Staubli VAL3: trajectory.pjx

--- trajectory.pjx ---
Parameters version=s8.15.3Cs9_BS3337 stackSize=5000 millimeterUnit=true
Program file=copy.pgx
Program file=copyPoint.pgx
Program file=copyPoint1.pgx
Program file=copyPoint3.pgx
Program file=deletePoint.pgx
Program file=deleteTraj.pgx
Program file=getFrameID.pgx
Program file=getIFvalue.pgx
Program file=getLibName.pgx
Program file=getMoveType.pgx
Program file=getPointIndex.pgx
Program file=getPointPara.pgx
Program file=getPointSize.pgx
Program file=getSize.pgx
Program file=getToolID.pgx
Program file=getTrajList.pgx
Program file=getTrajSize.pgx
Program file=insertAction.pgx
Program file=insertCirclePoint.pgx
Program file=insertDelay.pgx
Program file=insertENDIF.pgx
Program file=insertIF.pgx
Program file=insertJoint.pgx
Program file=insertPoint.pgx
Program file=insertSignal.pgx
Program file=isDefine.pgx
Program file=isPointOK.pgx
Program file=isReachable.pgx
Program file=loadTRAJ.pgx
Program file=logicIF.pgx
Program file=makeTraj.pgx
Program file=modifyAll.pgx
Program file=modifyPara.pgx
Program file=new.pgx
Program file=onSave.pgx
Program file=pointEdit.pgx
Program file=pointEditValue.pgx
Program file=pointMove.pgx
Program file=pointMove1.pgx
Program file=pointToString.pgx
Program file=resetMark.pgx
Program file=resizeMark.pgx
Program file=setMark.pgx
Program file=start.pgx
Program file=stop.pgx
Program file=teachPoint.pgx
Program file=teachPoint1.pgx
Data file=trajectory.dtx
Library alias=savedata path=Disk://source/saveData/saveData.pjx
Library alias=io path=Disk://source/projectSource/io/io.pjx
Library alias=rs path=Disk://source/projectSource/robotStatus/robotStatus.pjx
Library alias=actData path=Disk://data/actionData/actionData.pjx
Library alias=action path=Disk://source/projectSource/Action/Action.pjx
Library alias=trajTemp path=Disk://source/template/trajTemp/trajTemp.pjx
Library alias=ar path=Disk://autoReturn/autoReturn.pjx
Type name=pointItem path=Disk://source/template/pointItem/pointItem.pjx
Type name=trajItem path=Disk://source/template/trajItem/trajItem.pjx

--- trajectory.dtx ---
mdesc mNomSpeed
frame fFrame = {fatherId=world[0]}
tool tTool = {fatherId=flange[0]}
mdesc mSim = {blend=off}
frame _fFrame = {fatherId=world[0]}
pointRx pGOTO = {fatherId=world[0]}
num nIndex[100]

--- start.pgx ---
program start()
begin
end

--- copy.pgx ---
public program copy(string x_sSource, string& x_sTarget, bool& x_bToSave)
  local num l_j
  local num l_i
begin
  trajTemp:tTrajItem[x_sTarget].nFrameIndex=trajTemp:tTrajItem[x_sSource].nFrameIndex
  trajTemp:tTrajItem[x_sTarget].nToolIndex=trajTemp:tTrajItem[x_sSource].nToolIndex
  trajTemp:tTrajItem[x_sTarget].nMoveID=trajTemp:tTrajItem[x_sSource].nMoveID
  trajTemp:tTrajItem[x_sTarget].sID=trajTemp:tTrajItem[x_sTarget].sID
  resize(trajTemp:tTrajItem[x_sTarget].pPointItem,1,size(trajTemp:tTrajItem[x_sSource].pPointItem))
  for l_i = 0 to size(trajTemp:tTrajItem[x_sSource].pPointItem)-1
    trajTemp:tTrajItem[x_sTarget].pPointItem[l_i].pParaItem.mMdesc=trajTemp:tTrajItem[x_sSource].pPointItem[l_i].pParaItem.mMdesc
    trajTemp:tTrajItem[x_sTarget].pPointItem[l_i].pParaItem.nMoveType=trajTemp:tTrajItem[x_sSource].pPointItem[l_i].pParaItem.nMoveType
    trajTemp:tTrajItem[x_sTarget].pPointItem[l_i].pPointRx=trajTemp:tTrajItem[x_sSource].pPointItem[l_i].pPointRx
    //2025.03.18 add mlc  2025.10.16 modify by liu zhengang
    trajTemp:tTrajItem[x_sTarget].pPointItem[l_i].pInter=trajTemp:tTrajItem[x_sSource].pPointItem[l_i].pInter
    trajTemp:tTrajItem[x_sTarget].pPointItem[l_i].jJointRx=trajTemp:tTrajItem[x_sSource].pPointItem[l_i].jJointRx
    for l_j = 0 to 0
      trajTemp:tTrajItem[x_sTarget].pPointItem[l_i].pParaItem.nActionIndex[l_j]=trajTemp:tTrajItem[x_sSource].pPointItem[l_i].pParaItem.nActionIndex[l_j]
      trajTemp:tTrajItem[x_sTarget].pPointItem[l_i].pParaItem.nPercentage[l_j]=trajTemp:tTrajItem[x_sSource].pPointItem[l_i].pParaItem.nPercentage[l_j]
      trajTemp:tTrajItem[x_sTarget].pPointItem[l_i].pParaItem.iIfItem.bANDOR[l_j]=(trajTemp:tTrajItem[x_sSource].pPointItem[l_i].pParaItem.iIfItem.bANDOR[l_j]==true)
    endFor
    for l_j = 0 to 2
      trajTemp:tTrajItem[x_sTarget].pPointItem[l_i].pParaItem.iIfItem.nSigType[l_j]=trajTemp:tTrajItem[x_sSource].pPointItem[l_i].pParaItem.iIfItem.nSigType[l_j]
      trajTemp:tTrajItem[x_sTarget].pPointItem[l_i].pParaItem.iIfItem.nSigIndex[l_j]=trajTemp:tTrajItem[x_sSource].pPointItem[l_i].pParaItem.iIfItem.nSigIndex[l_j]
      trajTemp:tTrajItem[x_sTarget].pPointItem[l_i].pParaItem.iIfItem.nValue[l_j]=trajTemp:tTrajItem[x_sSource].pPointItem[l_i].pParaItem.iIfItem.nValue[l_j]
    endFor
    //
    trajTemp:tTrajItem[x_sTarget].pPointItem[l_i].pParaItem.nDelay=trajTemp:tTrajItem[x_sSource].pPointItem[l_i].pParaItem.nDelay
    trajTemp:tTrajItem[x_sTarget].pPointItem[l_i].pParaItem.nSigValue=trajTemp:tTrajItem[x_sSource].pPointItem[l_i].pParaItem.nSigValue
  endFor
  x_bToSave=true
end

--- copyPoint.pgx ---
public program copyPoint(string x_sKey, bool& x_bMark)
  local num l_nSize
  local num l_j
  local num l_i
begin
  resize(savedata:nMarkIndex,1,1)
  savedata:nMarkIndex=-1
  call getPointSize(x_sKey,l_nSize)
  l_j = 0
  for l_i = 0 to l_nSize-1
    if trajTemp:tTrajItem[x_sKey].pPointItem[l_i].bMarked
      l_j=l_j+1
      insert(savedata:nMarkIndex[l_j])
      savedata:nMarkIndex[l_j]=l_i


    endIf
  endFor
  x_bMark=false
end

--- copyPoint1.pgx ---
public program copyPoint1(string x_sKey, num x_nIndex)
  local num l_i
begin
  for l_i = 1 to size(savedata:nMarkIndex)-1
    insert(trajTemp:tTrajItem[x_sKey].pPointItem[x_nIndex+l_i])
    call copyPoint3(x_sKey,x_nIndex+l_i,savedata:nMarkIndex[l_i])
  endFor
  call resetMark(x_sKey)
end

--- copyPoint3.pgx ---
public program copyPoint3(string x_sKey, num x_nTarget, num x_nSource)
  local num l_i
begin
  trajTemp:tTrajItem[x_sKey].pPointItem[x_nTarget].pPointRx=trajTemp:tTrajItem[x_sKey].pPointItem[x_nSource].pPointRx
  //trajTemp:tTrajItem[x_sKey].pPointItem[x_nTarget].pPointRx[1]=trajTemp:tTrajItem[x_sKey].pPointItem[x_nSource].pPointRx[1]
  trajTemp:tTrajItem[x_sKey].pPointItem[x_nTarget].jJointRx=trajTemp:tTrajItem[x_sKey].pPointItem[x_nSource].jJointRx
  trajTemp:tTrajItem[x_sKey].pPointItem[x_nTarget].sID=trajTemp:tTrajItem[x_sKey].pPointItem[x_nSource].sID
  trajTemp:tTrajItem[x_sKey].pPointItem[x_nTarget].bMarked=trajTemp:tTrajItem[x_sKey].pPointItem[x_nSource].bMarked
  trajTemp:tTrajItem[x_sKey].pPointItem[x_nTarget].pInter=trajTemp:tTrajItem[x_sKey].pPointItem[x_nSource].pInter
  trajTemp:tTrajItem[x_sKey].pPointItem[x_nTarget].pParaItem.mMdesc=trajTemp:tTrajItem[x_sKey].pPointItem[x_nSource].pParaItem.mMdesc
  trajTemp:tTrajItem[x_sKey].pPointItem[x_nTarget].pParaItem.nMoveType=trajTemp:tTrajItem[x_sKey].pPointItem[x_nSource].pParaItem.nMoveType
  trajTemp:tTrajItem[x_sKey].pPointItem[x_nTarget].pParaItem.nActionIndex=trajTemp:tTrajItem[x_sKey].pPointItem[x_nSource].pParaItem.nActionIndex
  trajTemp:tTrajItem[x_sKey].pPointItem[x_nTarget].pParaItem.nPercentage=trajTemp:tTrajItem[x_sKey].pPointItem[x_nSource].pParaItem.nPercentage
  trajTemp:tTrajItem[x_sKey].pPointItem[x_nTarget].pParaItem.nDelay=trajTemp:tTrajItem[x_sKey].pPointItem[x_nSource].pParaItem.nDelay
  trajTemp:tTrajItem[x_sKey].pPointItem[x_nTarget].pParaItem.nSigValue=trajTemp:tTrajItem[x_sKey].pPointItem[x_nSource].pParaItem.nSigValue
  trajTemp:tTrajItem[x_sKey].pPointItem[x_nTarget].pParaItem.bSafePoint=trajTemp:tTrajItem[x_sKey].pPointItem[x_nSource].pParaItem.bSafePoint
  for l_i = 0 to 2
    trajTemp:tTrajItem[x_sKey].pPointItem[x_nTarget].pParaItem.iIfItem.nSigType[l_i]=trajTemp:tTrajItem[x_sKey].pPointItem[x_nSource].pParaItem.iIfItem.nSigType[l_i]
    trajTemp:tTrajItem[x_sKey].pPointItem[x_nTarget].pParaItem.iIfItem.nSigIndex[l_i]=trajTemp:tTrajItem[x_sKey].pPointItem[x_nSource].pParaItem.iIfItem.nSigIndex[l_i]
    trajTemp:tTrajItem[x_sKey].pPointItem[x_nTarget].pParaItem.iIfItem.nValue[l_i]=trajTemp:tTrajItem[x_sKey].pPointItem[x_nSource].pParaItem.iIfItem.nValue[l_i]
  endFor
  trajTemp:tTrajItem[x_sKey].pPointItem[x_nTarget].pParaItem.iIfItem.bANDOR[0]=trajTemp:tTrajItem[x_sKey].pPointItem[x_nSource].pParaItem.iIfItem.bANDOR[0]
  trajTemp:tTrajItem[x_sKey].pPointItem[x_nTarget].pParaItem.iIfItem.bANDOR[1]=trajTemp:tTrajItem[x_sKey].pPointItem[x_nSource].pParaItem.iIfItem.bANDOR[1]

end

--- deletePoint.pgx ---
public program deletePoint(string x_sKey, num x_nIndex, bool& x_bToSave)
  local bool l_bResult
begin
  l_bResult=userPageConfirm("是否删除点位："+toString("",x_nIndex))
  if l_bResult
    if x_nIndex==0 and size(trajTemp:tTrajItem[x_sKey].pPointItem)==1
      userPageAlert("数组元素不得为0")
    else
      delete(trajTemp:tTrajItem[x_sKey].pPointItem[x_nIndex])
      //trajTemp:libSave()
      x_bToSave=true
    endIf
  endIf

end

--- deleteTraj.pgx ---
public program deleteTraj(string x_sKey, bool& x_bToSave)
begin
  if isDefined(trajTemp:tTrajItem[x_sKey])
    delete(trajTemp:tTrajItem[x_sKey])
    //trajTemp:libSave()
  endIf
  x_bToSave=true
end

--- getFrameID.pgx ---
public program getFrameID(string x_sKey, num& x_nFrameID)
begin
  x_nFrameID=trajTemp:tTrajItem[x_sKey].nFrameIndex
end

--- getIFvalue.pgx ---
public program getIFvalue(string x_sKey, num x_nIndex, bool& x_bFinalResult)
  local num l_nSigType[3]
  local num l_i
  local num l_nSigValue[3]
  local bool l_bANDOR[2]
  local num l_nSigIndex[3]
  local bool l_bValue
  local bool l_bErr
  local bool l_bSetValue
  local num l_nResult[3]
  local bool l_bResult0[2]
  local num l_nValue
begin
  //l_nResult=0,null
  //         =1,true
  //         =2,false

  for l_i = 0 to 2
    l_nSigType[l_i]= trajTemp:tTrajItem[x_sKey].pPointItem[x_nIndex].pParaItem.iIfItem.nSigType[l_i]
    l_nSigValue[l_i]=trajTemp:tTrajItem[x_sKey].pPointItem[x_nIndex].pParaItem.iIfItem.nValue[l_i]
    l_nSigIndex[l_i]=trajTemp:tTrajItem[x_sKey].pPointItem[x_nIndex].pParaItem.iIfItem.nSigIndex[l_i]
  endFor
  l_bANDOR[0]=trajTemp:tTrajItem[x_sKey].pPointItem[x_nIndex].pParaItem.iIfItem.bANDOR[0]
  l_bANDOR[1]=trajTemp:tTrajItem[x_sKey].pPointItem[x_nIndex].pParaItem.iIfItem.bANDOR[1]

  for l_i = 0 to 2
    if l_nSigType[l_i]!=0 and l_nSigIndex[l_i]!=0
      switch l_nSigType[l_i]
        case 1
          //din
          call io:getDigIO(io:dInput[l_nSigIndex[l_i]],l_bValue,l_bErr)
          l_bSetValue=(l_nSigValue[l_i]!=0)
          if l_bSetValue==l_bValue
            l_nResult[l_i]=1
          else
            l_nResult[l_i]=2
          endIf
        break
        case 2
          //dout
          call io:getDigIO(io:dOutput[l_nSigIndex[l_i]],l_bValue,l_bErr)
          l_bSetValue=(l_nSigValue[l_i]!=0)
          if l_bSetValue==l_bValue
            l_nResult[l_i]=1
          else
            l_nResult[l_i]=2
          endIf
        break
        case 3
          //ain
          call io:getAnaIO(io:aInput[l_nSigIndex[l_i]],l_nValue,l_bErr)
          if l_nSigValue[l_i]==l_nValue
            l_nResult[l_i]=1
          else
            l_nResult[l_i]=2
          endIf
        break
        case 4
          //aout
          call io:getAnaIO(io:aOutput[l_nSigIndex[l_i]],l_nValue,l_bErr)
          if l_nSigValue[l_i]==l_nValue
            l_nResult[l_i]=1
          else
            l_nResult[l_i]=2
          endIf
        break
      endSwitch
    else
      l_nResult[l_i]=0
    endIf
  endFor

  //logic
 call logicIF(l_nResult[0],l_nResult[1],l_nResult[2],l_bANDOR[0],l_bANDOR[1],x_bFinalResult)

end

--- getLibName.pgx ---
public program getLibName(num& x_nLibNum, bool& x_bResult)
  local string l_sString
  local string l_sString1
  local num l_nPos
  local string l_sPath
  local num l_nlength
  local num l_nlength1
  local num l_nLength2
  local num l_nSize
  local string l_sTarget
  local num l_nLength
begin
  l_sPath=trajTemp:libPath()
  l_nlength=len("Disk://data/CustomerLib/lib")
  l_nlength1=len("/saveTRAJ/saveTRAJ.pjx")
  l_nLength2=len(l_sPath)
  l_nSize=l_nLength2-l_nlength1-l_nLength
  l_sTarget=mid(l_sPath,l_nSize,l_nlength)
  toNum(l_sTarget,x_nLibNum,x_bResult)
end

--- getMoveType.pgx ---
public program getMoveType(string x_sKey, num x_nIndex, num& x_nMoveType)
begin
  x_nMoveType=trajTemp:tTrajItem[x_sKey].pPointItem[x_nIndex].pParaItem.nMoveType
end

--- getPointIndex.pgx ---
public program getPointIndex(string x_sTrajItem, string x_sPoint, num& x_nPointIndex, bool& x_bResult)
  local bool l_bResult
  local num l_nSize
begin
  toNum(x_sPoint,x_nPointIndex,x_bResult)
  if !x_bResult
    call getPointSize(x_sTrajItem,l_nSize)
    x_nPointIndex=l_nSize-1
  endIf
end

--- getPointPara.pgx ---
public program getPointPara(string x_sKey, num x_nIndex, num& x_nMoveType, num& x_nParaSpeed, num& x_nParaAccel, num& x_nParaBlend, num x_nParaPercent, string& x_sComment, bool& x_bSafePoint, string& x_sBlend, num& x_nValue[], string& x_sTRSF[])
  local num l_nMoveType
begin
  x_nMoveType=trajTemp:tTrajItem[x_sKey].pPointItem[x_nIndex].pParaItem.nMoveType
  x_nParaSpeed=trajTemp:tTrajItem[x_sKey].pPointItem[x_nIndex].pParaItem.mMdesc.vel
  x_nParaAccel=trajTemp:tTrajItem[x_sKey].pPointItem[x_nIndex].pParaItem.mMdesc.accel
  x_nParaBlend=trajTemp:tTrajItem[x_sKey].pPointItem[x_nIndex].pParaItem.mMdesc.leave
  x_nParaPercent=trajTemp:tTrajItem[x_sKey].pPointItem[x_nIndex].pParaItem.nPercentage
  x_sComment=trajTemp:tTrajItem[x_sKey].pPointItem[x_nIndex].sID
  //  x_bBlendJoint=(trajTemp:tTrajItem[x_sKey].pPointItem[x_nIndex].pParaItem.mMdesc.blend==joint)
  //  x_bBlendOFF=(trajTemp:tTrajItem[x_sKey].pPointItem[x_nIndex].pParaItem.mMdesc.blend==off)
  switch x_nMoveType
    case 1

      x_nValue[0]=trajTemp:tTrajItem[x_sKey].pPointItem[x_nIndex].jJointRx.j1
      x_nValue[1]=trajTemp:tTrajItem[x_sKey].pPointItem[x_nIndex].jJointRx.j2
      x_nValue[2]=trajTemp:tTrajItem[x_sKey].pPointItem[x_nIndex].jJointRx.j3
      x_nValue[3]=trajTemp:tTrajItem[x_sKey].pPointItem[x_nIndex].jJointRx.j4
      x_nValue[4]=trajTemp:tTrajItem[x_sKey].pPointItem[x_nIndex].jJointRx.j5
      x_nValue[5]=trajTemp:tTrajItem[x_sKey].pPointItem[x_nIndex].jJointRx.j6

      x_sTRSF[0]="J1:"
      x_sTRSF[1]="J2:"
      x_sTRSF[2]="J3:"
      x_sTRSF[3]="J4:"
      x_sTRSF[4]="J5:"
      x_sTRSF[5]="J6:"

    break
    case 0
      x_nValue[0]=trajTemp:tTrajItem[x_sKey].pPointItem[x_nIndex].pPointRx.trsf.x
      x_nValue[1]=trajTemp:tTrajItem[x_sKey].pPointItem[x_nIndex].pPointRx.trsf.y
      x_nValue[2]=trajTemp:tTrajItem[x_sKey].pPointItem[x_nIndex].pPointRx.trsf.z
      x_nValue[3]=trajTemp:tTrajItem[x_sKey].pPointItem[x_nIndex].pPointRx.trsf.rx
      x_nValue[4]=trajTemp:tTrajItem[x_sKey].pPointItem[x_nIndex].pPointRx.trsf.ry
      x_nValue[5]=trajTemp:tTrajItem[x_sKey].pPointItem[x_nIndex].pPointRx.trsf.rz

      x_sTRSF[0]="X:"
      x_sTRSF[1]="Y:"
      x_sTRSF[2]="Z:"
      x_sTRSF[3]="RX:"
      x_sTRSF[4]="RY:"
      x_sTRSF[5]="RZ:"
    break
    case 2
      x_nValue[0]=trajTemp:tTrajItem[x_sKey].pPointItem[x_nIndex].pPointRx.trsf.x
      x_nValue[1]=trajTemp:tTrajItem[x_sKey].pPointItem[x_nIndex].pPointRx.trsf.y
      x_nValue[2]=trajTemp:tTrajItem[x_sKey].pPointItem[x_nIndex].pPointRx.trsf.z
      x_nValue[3]=trajTemp:tTrajItem[x_sKey].pPointItem[x_nIndex].pPointRx.trsf.rx
      x_nValue[4]=trajTemp:tTrajItem[x_sKey].pPointItem[x_nIndex].pPointRx.trsf.ry
      x_nValue[5]=trajTemp:tTrajItem[x_sKey].pPointItem[x_nIndex].pPointRx.trsf.rz
      x_nValue[6]= trajTemp:tTrajItem[x_sKey].pPointItem[x_nIndex].pInter.trsf.x
      x_nValue[7]=trajTemp:tTrajItem[x_sKey].pPointItem[x_nIndex].pInter.trsf.y
      x_nValue[8]=trajTemp:tTrajItem[x_sKey].pPointItem[x_nIndex].pInter.trsf.z
      x_nValue[9]=trajTemp:tTrajItem[x_sKey].pPointItem[x_nIndex].pInter.trsf.rx
      x_nValue[10]=trajTemp:tTrajItem[x_sKey].pPointItem[x_nIndex].pInter.trsf.ry
      x_nValue[11]= trajTemp:tTrajItem[x_sKey].pPointItem[x_nIndex].pInter.trsf.rz
      x_sTRSF[0]="X:"
      x_sTRSF[1]="Y:"
      x_sTRSF[2]="Z:"
      x_sTRSF[3]="RX:"
      x_sTRSF[4]="RY:"
      x_sTRSF[5]="RZ:"
      x_sTRSF[6]="2X:"
      x_sTRSF[7]="2Y:"
      x_sTRSF[8]="2Z:"
      x_sTRSF[9]="2RX:"
      x_sTRSF[10]="2RY:"
      x_sTRSF[11]="2RZ:"

    break
  endSwitch
  //blend
  if trajTemp:tTrajItem[x_sKey].pPointItem[x_nIndex].pParaItem.mMdesc.blend==off
    x_sBlend="OFF"
  elseIf trajTemp:tTrajItem[x_sKey].pPointItem[x_nIndex].pParaItem.mMdesc.blend==joint
    x_sBlend="关节"
  elseIf trajTemp:tTrajItem[x_sKey].pPointItem[x_nIndex].pParaItem.mMdesc.blend==Cartesian
    x_sBlend="笛卡尔"
  endIf
  x_bSafePoint = (trajTemp:tTrajItem[x_sKey].pPointItem.pParaItem.bSafePoint==true)
end

--- getPointSize.pgx ---
public program getPointSize(string x_sKey, num& x_nSize)
begin
  x_nSize=size(trajTemp:tTrajItem[x_sKey].pPointItem)
end

--- getSize.pgx ---
public program getSize(num& x_nSize)
begin
  if size(trajTemp:tTrajItem)>0
    x_nSize=size(trajTemp:tTrajItem)
  else
    x_nSize=0
  endIf
end

--- getToolID.pgx ---
public program getToolID(string x_sKey, num& x_nToolID)
begin
   x_nToolID=trajTemp:tTrajItem[x_sKey].nToolIndex
end

--- getTrajList.pgx ---
public program getTrajList(string& x_sList[])
  local string l_sKey
begin
  resize(x_sList,1,1)
  l_sKey=first(trajTemp:tTrajItem)

  while l_sKey!=""
    x_sList[size(x_sList)-1]=l_sKey

    l_sKey=next(trajTemp:tTrajItem[l_sKey])

    if l_sKey!=""
      insert(x_sList[size(x_sList)])
    endIf
  endWhile
  if size(trajTemp:tTrajItem)<1
    x_sList=""
  endIf
end

--- getTrajSize.pgx ---
public program getTrajSize(num& x_nSize)
begin
  x_nSize=size(trajTemp:tTrajItem)
end

--- insertAction.pgx ---
public program insertAction(string x_sKey, num x_nIndex, num x_nValue, bool& x_bToSave)
  local num l_i
begin
  // insert(trajTemp:tTrajItem[x_sKey].pPointItem[x_nIndex+1])
  append(trajTemp:tTrajItem[x_sKey].pPointItem)

  for l_i = (size(trajTemp:tTrajItem[x_sKey].pPointItem)-1) to(x_nIndex+1) step -1
    //logMsg(toString("",l_i))
    call copyPoint3(x_sKey,l_i,l_i-1)
  endFor
  trajTemp:tTrajItem[x_sKey].pPointItem[x_nIndex+1].pParaItem.nMoveType=10
  trajTemp:tTrajItem[x_sKey].pPointItem[x_nIndex+1].pParaItem.nSigValue=x_nValue
  //trajTemp:libSave()
  x_bToSave=true
end

--- insertCirclePoint.pgx ---
public program insertCirclePoint(string x_sKey, num x_nIndex, bool& x_bToSave)
  local num l_j
  local frame l_fFrame
  local tool l_tTool
  local num l_i
  local num l_nFrameIndex
  local num l_nToolIndex
  local pointRx l_pPoint
begin
  //  link(l_fFrame,world)
  //  link(l_tTool,flange)
  //  call savedata:getFrame(trajTemp:tTrajItem[x_sKey].nFrameIndex,l_fFrame)
  //  call savedata:getTool(trajTemp:tTrajItem[x_sKey].nToolIndex,l_tTool)
  //insert(trajTemp:tTrajItem[x_sKey].pPointItem[x_nIndex+1])
  append(trajTemp:tTrajItem[x_sKey].pPointItem)

  for l_i = (size(trajTemp:tTrajItem[x_sKey].pPointItem)-1) to(x_nIndex+1) step -1
    //logMsg(toString("",l_i))
    call copyPoint3(x_sKey,l_i,l_i-1)
  endFor
  //2024.12.06 当前位置作为插入点坐标
  l_nFrameIndex=trajTemp:tTrajItem[x_sKey].nFrameIndex
  l_nToolIndex=trajTemp:tTrajItem[x_sKey].nToolIndex
  call savedata:getFrame(l_nFrameIndex,l_fFrame)
  call savedata:getTool(l_nToolIndex,l_tTool)
  trajTemp:tTrajItem[x_sKey].pPointItem[x_nIndex+1].jJointRx=herej()
  l_pPoint=jointToPoint(l_tTool,l_fFrame,herej())
  trajTemp:tTrajItem[x_sKey].pPointItem[x_nIndex+1].pPointRx.trsf=l_pPoint.trsf
  trajTemp:tTrajItem[x_sKey].pPointItem[x_nIndex+1].pPointRx.config=l_pPoint.config
  trajTemp:tTrajItem[x_sKey].pPointItem[x_nIndex+1].pInter.trsf=l_pPoint.trsf
  trajTemp:tTrajItem[x_sKey].pPointItem[x_nIndex+1].pInter.config=l_pPoint.config
  //

  //trajTemp:tTrajItem[x_sKey].pPointItem[x_nIndex+1].pPointRx=trajTemp:tTrajItem[x_sKey].pPointItem[x_nIndex].pPointRx
  //trajTemp:tTrajItem[x_sKey].pPointItem[x_nIndex+1].jJointRx=trajTemp:tTrajItem[x_sKey].pPointItem[x_nIndex].jJointRx
  trajTemp:tTrajItem[x_sKey].pPointItem[x_nIndex+1].pParaItem.mMdesc=trajTemp:tTrajItem[x_sKey].pPointItem[x_nIndex].pParaItem.mMdesc
  trajTemp:tTrajItem[x_sKey].pPointItem[x_nIndex+1].pParaItem.nMoveType=2
  trajTemp:tTrajItem[x_sKey].pPointItem[x_nIndex+1].pParaItem.nDelay=trajTemp:tTrajItem[x_sKey].pPointItem[x_nIndex].pParaItem.nDelay
  trajTemp:tTrajItem[x_sKey].pPointItem[x_nIndex+1].pParaItem.nSigValue=trajTemp:tTrajItem[x_sKey].pPointItem[x_nIndex].pParaItem.nSigValue
  trajTemp:tTrajItem[x_sKey].pPointItem[x_nIndex+1].pParaItem.nActionIndex=trajTemp:tTrajItem[x_sKey].pPointItem[x_nIndex].pParaItem.nActionIndex
  trajTemp:tTrajItem[x_sKey].pPointItem[x_nIndex+1].pParaItem.nPercentage=trajTemp:tTrajItem[x_sKey].pPointItem[x_nIndex].pParaItem.nPercentage
  for l_j = 0 to 2
    trajTemp:tTrajItem[x_sKey].pPointItem[x_nIndex+1].pParaItem.iIfItem.nSigType[l_j]=trajTemp:tTrajItem[x_sKey].pPointItem[x_nIndex].pParaItem.iIfItem.nSigType[l_j]
    trajTemp:tTrajItem[x_sKey].pPointItem[x_nIndex+1].pParaItem.iIfItem.nSigIndex[l_j]=trajTemp:tTrajItem[x_sKey].pPointItem[x_nIndex].pParaItem.iIfItem.nSigIndex[l_j]
    trajTemp:tTrajItem[x_sKey].pPointItem[x_nIndex+1].pParaItem.iIfItem.nValue[l_j]=trajTemp:tTrajItem[x_sKey].pPointItem[x_nIndex].pParaItem.iIfItem.nValue[l_j]
  endFor
  //trajTemp:libSave()
  x_bToSave=true
end

--- insertDelay.pgx ---
public program insertDelay(string x_sKey, num x_nIndex, bool& x_bToSave, num x_nMoveType, num x_nDelay)
  local num l_j
  local num l_i
begin
  //insert(trajTemp:tTrajItem[x_sKey].pPointItem[x_nIndex+1])
  append(trajTemp:tTrajItem[x_sKey].pPointItem)

  for l_i = (size(trajTemp:tTrajItem[x_sKey].pPointItem)-1) to(x_nIndex+1) step -1
   // logMsg(toString("",l_i))
    call copyPoint3(x_sKey,l_i,l_i-1)
  endFor
  trajTemp:tTrajItem[x_sKey].pPointItem[x_nIndex+1].pParaItem.nMoveType=x_nMoveType

  trajTemp:tTrajItem[x_sKey].pPointItem[x_nIndex+1].pParaItem.nDelay=x_nDelay

 //trajTemp:libSave()

  x_bToSave=true
end

--- insertENDIF.pgx ---
public program insertENDIF(string x_sKey, num x_nIndex, bool& x_bToSave)
  local num l_j
  local num l_i
begin

  //insert(trajTemp:tTrajItem[x_sKey].pPointItem[x_nIndex+1])
  append(trajTemp:tTrajItem[x_sKey].pPointItem)

  for l_i = (size(trajTemp:tTrajItem[x_sKey].pPointItem)-1) to(x_nIndex+1) step -1
    //logMsg(toString("",l_i))
    call copyPoint3(x_sKey,l_i,l_i-1)
  endFor
  trajTemp:tTrajItem[x_sKey].pPointItem[x_nIndex+1].pParaItem.nMoveType=9

  //trajTemp:libSave()
  x_bToSave=true
end

--- insertIF.pgx ---
public program insertIF(string x_sKey, num x_nIndex, num& x_nMoveType[], num& x_nIOIndex[], num& x_nValue[], num& x_nANDOR[], bool& x_bToSave)
  local num l_j
  local num l_i
begin
  // insert(trajTemp:tTrajItem[x_sKey].pPointItem[x_nIndex+1])
  append(trajTemp:tTrajItem[x_sKey].pPointItem)

  for l_i = (size(trajTemp:tTrajItem[x_sKey].pPointItem)-1) to(x_nIndex+1) step -1
    // logMsg(toString("",l_i))
    call copyPoint3(x_sKey,l_i,l_i-1)
  endFor
  trajTemp:tTrajItem[x_sKey].pPointItem[x_nIndex+1].pParaItem.nMoveType=8
  for l_i =0 to 2
    trajTemp:tTrajItem[x_sKey].pPointItem[x_nIndex+1].pParaItem.iIfItem.nSigType[l_i]=x_nMoveType[l_i]
    trajTemp:tTrajItem[x_sKey].pPointItem[x_nIndex+1].pParaItem.iIfItem.nSigIndex[l_i]=x_nIOIndex[l_i]
    trajTemp:tTrajItem[x_sKey].pPointItem[x_nIndex+1].pParaItem.iIfItem.nValue[l_i]=x_nValue[l_i]
  endFor
  for l_i = 0 to 1
    trajTemp:tTrajItem[x_sKey].pPointItem[x_nIndex+1].pParaItem.iIfItem.bANDOR[l_i]=(x_nANDOR[l_i]==2)
  endFor

  //trajTemp:libSave()
  x_bToSave=true
end

--- insertJoint.pgx ---
public program insertJoint(string x_sKey, num x_nIndex, bool& x_bToSave)
  local num l_j
  local num l_i
begin
  // insert(trajTemp:tTrajItem[x_sKey].pPointItem[x_nIndex+1])
  append(trajTemp:tTrajItem[x_sKey].pPointItem)

  for l_i = (size(trajTemp:tTrajItem[x_sKey].pPointItem)-1) to(x_nIndex+1) step -1
    //logMsg(toString("",l_i))
    call copyPoint3(x_sKey,l_i,l_i-1)
  endFor
  trajTemp:tTrajItem[x_sKey].pPointItem[x_nIndex+1].pPointRx=trajTemp:tTrajItem[x_sKey].pPointItem[x_nIndex].pPointRx
  trajTemp:tTrajItem[x_sKey].pPointItem[x_nIndex+1].jJointRx=trajTemp:tTrajItem[x_sKey].pPointItem[x_nIndex].jJointRx
  trajTemp:tTrajItem[x_sKey].pPointItem[x_nIndex+1].pParaItem.mMdesc=trajTemp:tTrajItem[x_sKey].pPointItem[x_nIndex].pParaItem.mMdesc
  trajTemp:tTrajItem[x_sKey].pPointItem[x_nIndex+1].pParaItem.nMoveType=0
  trajTemp:tTrajItem[x_sKey].pPointItem[x_nIndex+1].pParaItem.nDelay=trajTemp:tTrajItem[x_sKey].pPointItem[x_nIndex].pParaItem.nDelay
  trajTemp:tTrajItem[x_sKey].pPointItem[x_nIndex+1].pParaItem.nSigValue=trajTemp:tTrajItem[x_sKey].pPointItem[x_nIndex].pParaItem.nSigValue
  trajTemp:tTrajItem[x_sKey].pPointItem[x_nIndex+1].pParaItem.nActionIndex=trajTemp:tTrajItem[x_sKey].pPointItem[x_nIndex].pParaItem.nActionIndex
  trajTemp:tTrajItem[x_sKey].pPointItem[x_nIndex+1].pParaItem.nPercentage=trajTemp:tTrajItem[x_sKey].pPointItem[x_nIndex].pParaItem.nPercentage
  for l_j = 0 to 2
    trajTemp:tTrajItem[x_sKey].pPointItem[x_nIndex+1].pParaItem.iIfItem.nSigType[l_j]=trajTemp:tTrajItem[x_sKey].pPointItem[x_nIndex].pParaItem.iIfItem.nSigType[l_j]
    trajTemp:tTrajItem[x_sKey].pPointItem[x_nIndex+1].pParaItem.iIfItem.nSigIndex[l_j]=trajTemp:tTrajItem[x_sKey].pPointItem[x_nIndex].pParaItem.iIfItem.nSigIndex[l_j]
    trajTemp:tTrajItem[x_sKey].pPointItem[x_nIndex+1].pParaItem.iIfItem.nValue[l_j]=trajTemp:tTrajItem[x_sKey].pPointItem[x_nIndex].pParaItem.iIfItem.nValue[l_j]
  endFor
  //trajTemp:libSave()
  x_bToSave=true
end

--- insertPoint.pgx ---
public program insertPoint(string x_sKey, num x_nIndex, bool& x_bToSave)
  local num l_j
  local frame l_fFrame
  local tool l_tTool
  local num l_i
begin
  //  link(l_fFrame,world)
  //  link(l_tTool,flange)
  //  call savedata:getFrame(trajTemp:tTrajItem[x_sKey].nFrameIndex,l_fFrame)
  //  call savedata:getTool(trajTemp:tTrajItem[x_sKey].nToolIndex,l_tTool)
  //insert(trajTemp:tTrajItem[x_sKey].pPointItem[x_nIndex+1])
   append(trajTemp:tTrajItem[x_sKey].pPointItem)

  for l_i = (size(trajTemp:tTrajItem[x_sKey].pPointItem)-1) to(x_nIndex+1) step -1
    //logMsg(toString("",l_i))
    call copyPoint3(x_sKey,l_i,l_i-1)
  endFor
  trajTemp:tTrajItem[x_sKey].pPointItem[x_nIndex+1].pPointRx=trajTemp:tTrajItem[x_sKey].pPointItem[x_nIndex].pPointRx
  trajTemp:tTrajItem[x_sKey].pPointItem[x_nIndex+1].jJointRx=trajTemp:tTrajItem[x_sKey].pPointItem[x_nIndex].jJointRx
  trajTemp:tTrajItem[x_sKey].pPointItem[x_nIndex+1].pParaItem.mMdesc=trajTemp:tTrajItem[x_sKey].pPointItem[x_nIndex].pParaItem.mMdesc
  trajTemp:tTrajItem[x_sKey].pPointItem[x_nIndex+1].pParaItem.nMoveType=1
  trajTemp:tTrajItem[x_sKey].pPointItem[x_nIndex+1].pParaItem.nDelay=trajTemp:tTrajItem[x_sKey].pPointItem[x_nIndex].pParaItem.nDelay
  trajTemp:tTrajItem[x_sKey].pPointItem[x_nIndex+1].pParaItem.nSigValue=trajTemp:tTrajItem[x_sKey].pPointItem[x_nIndex].pParaItem.nSigValue
  trajTemp:tTrajItem[x_sKey].pPointItem[x_nIndex+1].pParaItem.nActionIndex=trajTemp:tTrajItem[x_sKey].pPointItem[x_nIndex].pParaItem.nActionIndex
  trajTemp:tTrajItem[x_sKey].pPointItem[x_nIndex+1].pParaItem.nPercentage=trajTemp:tTrajItem[x_sKey].pPointItem[x_nIndex].pParaItem.nPercentage
  for l_j = 0 to 2
    trajTemp:tTrajItem[x_sKey].pPointItem[x_nIndex+1].pParaItem.iIfItem.nSigType[l_j]=trajTemp:tTrajItem[x_sKey].pPointItem[x_nIndex].pParaItem.iIfItem.nSigType[l_j]
    trajTemp:tTrajItem[x_sKey].pPointItem[x_nIndex+1].pParaItem.iIfItem.nSigIndex[l_j]=trajTemp:tTrajItem[x_sKey].pPointItem[x_nIndex].pParaItem.iIfItem.nSigIndex[l_j]
    trajTemp:tTrajItem[x_sKey].pPointItem[x_nIndex+1].pParaItem.iIfItem.nValue[l_j]=trajTemp:tTrajItem[x_sKey].pPointItem[x_nIndex].pParaItem.iIfItem.nValue[l_j]
  endFor
  //trajTemp:libSave()
  x_bToSave=true
end

--- insertSignal.pgx ---
public program insertSignal(string x_sKey, num x_nIndex, bool& x_bToSave, num x_nMoveType, num x_nActionIndex, num x_nSigValue)
  local num l_j
  local bool l_bResult
  local num l_nIndex
  local num l_i
begin
  l_nIndex=x_nIndex+1

  //insert(trajTemp:tTrajItem[x_sKey].pPointItem[l_nIndex])
  append(trajTemp:tTrajItem[x_sKey].pPointItem)

  for l_i = (size(trajTemp:tTrajItem[x_sKey].pPointItem)-1) to l_nIndex step -1
    // logMsg(toString("",l_i))
    call copyPoint3(x_sKey,l_i,l_i-1)
  endFor
  trajTemp:tTrajItem[x_sKey].pPointItem[l_nIndex].pParaItem.nMoveType=x_nMoveType

  trajTemp:tTrajItem[x_sKey].pPointItem[l_nIndex].pParaItem.nSigValue=x_nSigValue

  trajTemp:tTrajItem[x_sKey].pPointItem[l_nIndex].pParaItem.nActionIndex=x_nActionIndex



  x_bToSave=true
  //trajTemp:libSave()
end

--- isDefine.pgx ---
public program isDefine(string x_sKey, bool& x_bResult)
begin
  x_bResult=isDefined(trajTemp:tTrajItem[x_sKey])
end

--- isPointOK.pgx ---
public program isPointOK(string x_sKey, num x_nIndex, bool& x_bResult)
  local pointRx l_pPoint
  local num l_nToolID
  local tool l_tTool
  local frame l_fFrame
  local num l_nFrameID
  local bool l_bResult
  local jointRx l_jResult
begin
  link(l_tTool,flange)
  link(l_fFrame,world)
  call getFrameID(x_sKey,l_nFrameID)
  call getToolID(x_sKey,l_nToolID)
  call savedata:getTool(l_nToolID,l_tTool)
  call savedata:getFrame(l_nFrameID,l_fFrame)
  link(l_pPoint,l_fFrame)
  l_pPoint.trsf=trajTemp:tTrajItem[x_sKey].pPointItem[x_nIndex].pPointRx.trsf
  l_pPoint.config=trajTemp:tTrajItem[x_sKey].pPointItem[x_nIndex].pPointRx.config

  l_bResult=pointToJoint(l_tTool,herej(),l_pPoint,l_jResult)
  if l_pPoint.trsf!={0,0,0,0,0,0} and l_bResult and isInRange(l_jResult)
    x_bResult=true
  else
    x_bResult=false
  endIf
end

--- isReachable.pgx ---
public program isReachable(string x_sKey, num x_nIndex, tool x_tTool)
  local pointRx l_pPoint
  local bool l_bResult
  local mdesc l_mDesc
  local jointRx l_jJoint
begin
  if trajTemp:tTrajItem[x_sKey].pPointItem[x_nIndex].pParaItem.nMoveType==0
    l_mDesc=trajTemp:tTrajItem[x_sKey].pPointItem[x_nIndex].pParaItem.mMdesc
    l_pPoint.trsf=trajTemp:tTrajItem[x_sKey].pPointItem.pPointRx.trsf
    l_pPoint.config=trajTemp:tTrajItem[x_sKey].pPointItem.pPointRx.config
    l_bResult= pointToJoint(x_tTool,herej(),l_pPoint,l_jJoint)
    if l_bResult
      movel(l_pPoint,x_tTool,l_mDesc)
    endIf
  endIf
end

--- loadTRAJ.pgx ---
public program loadTRAJ(num x_nLib, num& x_nResult)
  local string l_sPath
  local num l_nResult
begin
  if x_nLib>=0
    l_sPath="Disk://data/CustomerLib/lib"+toString("",x_nLib)+"/saveTRAJ"
    //  if libList()
    //    endIf
    x_nResult=trajTemp:libLoad(l_sPath)
    if x_nResult!=0
      popUpMsg("2")
      call rs:setAlarm(300,0)
    endIf
  else
    call rs:setAlarm(302,0)
  endIf
end

--- logicIF.pgx ---
public program logicIF(num x_nResult1, num x_nResult2, num x_nResult3, bool x_bANDOR1, bool x_bANDOR2, bool& x_bFinalResult)
  local bool l_bFinalResult1
  local bool l_bFinalResult2
begin
  if x_nResult1==0 and x_nResult2==0 and x_nResult3==0
    x_bFinalResult=false
  elseIf x_nResult1==0 and x_nResult2==0 and x_nResult3!=0
    x_bFinalResult=(x_nResult3==1)
  elseIf x_nResult1==0 and x_nResult2!=0 and x_nResult3==0
    x_bFinalResult=(x_nResult2==1)
  elseIf x_nResult1!=0 and x_nResult2==0 and x_nResult3==0
    x_bFinalResult=(x_nResult1==1)
  elseIf x_nResult1!=0 and x_nResult2!=0 and x_nResult3==0
    if x_bANDOR1
      x_bFinalResult=(x_nResult1==1 or x_nResult2==1)
    else
      x_bFinalResult=(x_nResult1==1 and x_nResult2==1)
    endIf
  elseIf x_nResult1==0 and x_nResult2!=0 and x_nResult3!=0
    if x_bANDOR2
      x_bFinalResult=(x_nResult1==1 or x_nResult2==1)
    else
      x_bFinalResult=(x_nResult1==1 and x_nResult2==1)
    endIf
  elseIf x_nResult1!=0 and x_nResult2!=0 and x_nResult3!=0
    if x_bANDOR1 and x_bANDOR2
      x_bFinalResult=(x_nResult1==1 or x_nResult2==1 or x_nResult3==1)
    elseIf !x_bANDOR1 and !x_bANDOR2
      x_bFinalResult=(x_nResult1==1 and x_nResult2==1 and x_nResult3==1)
    elseIf !x_bANDOR1 and x_bANDOR2
      x_bFinalResult=(x_nResult1==1 and x_nResult2==1 or x_nResult3==1)
    elseIf x_bANDOR1 and !x_bANDOR2
      x_bFinalResult=((x_nResult1==1 or x_nResult2==1) and x_nResult3==1)
    endIf

  endIf
end

--- makeTraj.pgx ---
public program makeTraj(string x_sKey)
  local num l_nMoveType
  local num l_nMoveID
  local frame l_fFrame
  local tool l_tTool
  local pointRx l_pPoint[2]
  local jointRx l_jJoint
  local mdesc l_mDesc
  local num l_nSigIndex
  local num l_nValue
  local bool l_bErr
  local num l_nSigValue
  local bool l_bValue
  local bool l_bSigValue
  local num l_i
  local num l_nDelay
  local bool l_bResult
  local num l_nActIndex
  local num l_nGetID
  local string l_sMsg
begin
  rs:sTrajStatus="执行轨迹："+x_sKey
  rs:sCycleItem=x_sKey
  l_nMoveID=trajTemp:tTrajItem[x_sKey].nMoveID
  rs:nFrameIndex=trajTemp:tTrajItem[x_sKey].nFrameIndex
  rs:nToolIndex=trajTemp:tTrajItem[x_sKey].nToolIndex
  call savedata:getFrame(rs:nFrameIndex,l_fFrame)
  call savedata:getTool(rs:nToolIndex,l_tTool)
  waitEndMove()
  setMoveId(l_nMoveID)
  for l_i = 0 to size(trajTemp:tTrajItem[x_sKey].pPointItem)-1
    l_nMoveType=trajTemp:tTrajItem[x_sKey].pPointItem[l_i].pParaItem.nMoveType
    rs:nCycleIndex=l_i
    if !rs:bGOTO
      switch l_nMoveType
        case 1
          link(l_pPoint,l_fFrame)
          l_pPoint.trsf=trajTemp:tTrajItem[x_sKey].pPointItem[l_i].pPointRx.trsf
          l_pPoint.config=trajTemp:tTrajItem[x_sKey].pPointItem[l_i].pPointRx.config
          l_mDesc=trajTemp:tTrajItem[x_sKey].pPointItem[l_i].pParaItem.mMdesc
          //l_nGetID=movel(l_pPoint,l_tTool,l_mDesc)
          call ar:MoveL(l_pPoint,l_tTool,l_mDesc,l_nGetID,false)
          wait(getMoveId()>=l_nGetID)
          call pointToString(l_sMsg,x_sKey,l_i)
          //rs:sTrajStatus="移动到:"+toString("",l_i)+l_sMsg
          rs:sTrajStatus="["+x_sKey+"]移动到:"+toString("",l_i)+l_sMsg
        break
        case 0
          l_jJoint=trajTemp:tTrajItem[x_sKey].pPointItem[l_i].jJointRx
          l_mDesc=trajTemp:tTrajItem[x_sKey].pPointItem[l_i].pParaItem.mMdesc
          //l_nGetID=movej(l_jJoint,l_tTool,l_mDesc)
          call ar:MoveJ(l_jJoint,l_tTool,l_mDesc,l_nGetID,false)
          wait(getMoveId()>=l_nGetID)
          call pointToString(l_sMsg,x_sKey,l_i)
          //rs:sTrajStatus="移动到:"+toString("",l_i)+l_sMsg
          rs:sTrajStatus="["+x_sKey+"]移动到:"+toString("",l_i)+l_sMsg
        break
        case 2
          //2024.12.23 add 圆弧运动
          link(l_pPoint,l_fFrame)
          link(l_pPoint[1],l_fFrame)
          l_pPoint.trsf=trajTemp:tTrajItem[x_sKey].pPointItem[l_i].pInter.trsf
          l_pPoint.config=trajTemp:tTrajItem[x_sKey].pPointItem[l_i].pInter.config
          l_pPoint[1].trsf=trajTemp:tTrajItem[x_sKey].pPointItem[l_i].pPointRx.trsf
          l_pPoint[1].config=trajTemp:tTrajItem[x_sKey].pPointItem[l_i].pPointRx.config
          l_mDesc=trajTemp:tTrajItem[x_sKey].pPointItem[l_i].pParaItem.mMdesc
          //l_nGetID=movec(l_pPoint,l_pPoint[1],l_tTool,l_mDesc)
          call ar:MoveC(l_pPoint,l_pPoint[1],l_tTool,l_mDesc,l_nGetID)
          wait(getMoveId()>=l_nGetID)
          call pointToString(l_sMsg,x_sKey,l_i)
          //rs:sTrajStatus="移动到:"+toString("",l_i)+l_sMsg
          rs:sTrajStatus="["+x_sKey+"]移动到:"+toString("",l_i)+l_sMsg
        break
        case 3
          //dIn
          waitEndMove()
          l_nSigIndex=trajTemp:tTrajItem[x_sKey].pPointItem[l_i].pParaItem.nActionIndex
          l_bSigValue=(trajTemp:tTrajItem[x_sKey].pPointItem[l_i].pParaItem.nSigValue!=0)
          //call io:getDigIO(io:dInput[l_nSigIndex],l_bValue,l_bErr)
          call pointToString(l_sMsg,x_sKey,l_i)
          //rs:sTrajStatus="移动到:"+toString("",l_i)+l_sMsg
          rs:sTrajStatus="["+x_sKey+"]移动到:"+toString("",l_i)+l_sMsg
          // wait(l_bValue==l_bSigValue)
          call io:waitDigInput(io:dInput[l_nSigIndex],l_bSigValue,l_bErr)
        break
        case 4
          //dOut
          waitEndMove()
          l_nSigIndex=trajTemp:tTrajItem[x_sKey].pPointItem[l_i].pParaItem.nActionIndex
          l_bSigValue=(trajTemp:tTrajItem[x_sKey].pPointItem[l_i].pParaItem.nSigValue!=0)
          call io:setDigOutput(io:dOutput[l_nSigIndex],l_bSigValue,l_bErr)
          call pointToString(l_sMsg,x_sKey,l_i)
          //rs:sTrajStatus="移动到:"+toString("",l_i)+l_sMsg
          rs:sTrajStatus="["+x_sKey+"]移动到:"+toString("",l_i)+l_sMsg
        break
        case 5
          //ain
          waitEndMove()
          l_nSigIndex=trajTemp:tTrajItem[x_sKey].pPointItem[l_i].pParaItem.nActionIndex
          l_nSigValue=trajTemp:tTrajItem[x_sKey].pPointItem[l_i].pParaItem.nSigValue
          // call io:getAnaIO(io:aInput[l_nSigIndex],l_nValue,l_bErr)
          call pointToString(l_sMsg,x_sKey,l_i)
          //rs:sTrajStatus="移动到:"+toString("",l_i)+l_sMsg
          rs:sTrajStatus="["+x_sKey+"]移动到:"+toString("",l_i)+l_sMsg
          call io:waitAnaInput(io:aInput[l_nSigIndex],l_nSigValue,l_bErr)
          // wait(l_nSigValue==l_nValue)
        break
        case 6
          //aout
          waitEndMove()
          l_nSigIndex=trajTemp:tTrajItem[x_sKey].pPointItem[l_i].pParaItem.nActionIndex
          l_nSigValue=trajTemp:tTrajItem[x_sKey].pPointItem[l_i].pParaItem.nSigValue
          call io:setAnaOutput(io:aOutput[l_nSigIndex],l_nSigValue,l_bErr)
          call pointToString(l_sMsg,x_sKey,l_i)
          //rs:sTrajStatus="移动到:"+toString("",l_i)+l_sMsg
          rs:sTrajStatus="["+x_sKey+"]移动到:"+toString("",l_i)+l_sMsg
        break
        case 7
          //delay
          l_nDelay=trajTemp:tTrajItem[x_sKey].pPointItem[l_i].pParaItem.nDelay
          waitEndMove()
          call pointToString(l_sMsg,x_sKey,l_i)
          //rs:sTrajStatus="移动到:"+toString("",l_i)+l_sMsg
          rs:sTrajStatus="["+x_sKey+"]移动到:"+toString("",l_i)+l_sMsg
          delay(l_nDelay)
        break
        case 8
          //if
          waitEndMove()
          call getIFvalue(x_sKey,l_i,l_bResult)
          if l_bResult
            rs:sTrajStatus="IF条件满足，继续执行"
          else
            rs:sTrajStatus="IF条件不满足，跳过当前程序"
          endIf
          rs:bGOTO=(l_bResult==false)
        break
        case 9
          //endif
          rs:bGOTO=false
        break
        case 10
          rs:sTrajStatus="执行action->"+toString("",l_nActIndex)
          l_nActIndex=trajTemp:tTrajItem[x_sKey].pPointItem[l_i].pParaItem.nSigValue
          call action:action_do(l_nActIndex)
        break
        case 11
          //2025.7.21 add 喷淋delay
          call io:getAnaIO(io:aInput[3],l_nDelay,l_bErr)
          //l_nDelay=trajTemp:tTrajItem[x_sKey].pPointItem[l_i].pParaItem.nDelay
          waitEndMove()
          call pointToString(l_sMsg,x_sKey,l_i)
          rs:sTrajStatus="移动到轨迹"+x_sKey+":"+toString("",l_i)+l_sMsg
          delay(l_nDelay)
        break
//        case 12
//          waitEndMove()
//          //Axis1位置输出
//          call io:setDigOutput(io:dOutput[60],true,l_bErr)
//          l_nSigValue=trajTemp:tTrajItem[x_sKey].pPointItem[l_i].pParaItem.nSigValue
//          rs:sTrajStatus="移动L轴->"+toString("",l_nSigValue)
//          call io:setAnaOutput(io:aOutput[7],l_nSigValue,l_bErr)
//          //等待Axis1到位
//          call io:waitDigInput(io:dInput[60],true,l_bErr)
//          rs:sTrajStatus="等待L轴位置->"+toString("",l_nSigValue)+"到达"
//          //复位Axis1控制命令
//          call io:setDigOutput(io:dOutput[60],false,l_bErr)
//        break
//        case 13
//          waitEndMove()
//          //Axis2位置输出
//          call io:setDigOutput(io:dOutput[61],true,l_bErr)
//          l_nSigValue=trajTemp:tTrajItem[x_sKey].pPointItem[l_i].pParaItem.nSigValue
//          rs:sTrajStatus="移动R轴->"+toString("",l_nSigValue)
//          call io:setAnaOutput(io:aOutput[8],l_nSigValue,l_bErr)
//          //等待Axis2到位
//          call io:waitDigInput(io:dInput[61],true,l_bErr)
//          rs:sTrajStatus="等待R轴位置->"+toString("",l_nSigValue)+"到达"
//          //复位Axis2控制命令
//          call io:setDigOutput(io:dOutput[61],false,l_bErr)
//        break
//        case 14
//          waitEndMove()
//           //Axis3位置输出
//          call io:setDigOutput(io:dOutput[62],true,l_bErr)
//          l_nSigValue=trajTemp:tTrajItem[x_sKey].pPointItem[l_i].pParaItem.nSigValue
//          rs:sTrajStatus="移动Z轴->"+toString("",l_nSigValue)
//          call io:setAnaOutput(io:aOutput[9],l_nSigValue,l_bErr)
//          //等待Axis3到位
//          call io:waitDigInput(io:dInput[62],true,l_bErr)
//          rs:sTrajStatus="等待Z轴位置->"+toString("",l_nSigValue)+"到达"
//          //复位Axis3控制命令
//          call io:setDigOutput(io:dOutput[62],false,l_bErr)
//        break
      endSwitch
    else
      if l_nMoveType==9
        rs:bGOTO=false
      endIf
    endIf
    delay(0)
  endFor
  waitEndMove()
end

--- modifyAll.pgx ---
public program modifyAll(string x_sKey, num x_nMoveType, num x_nParaSpeed, num x_nParaBlend, num x_nParaPercent, string x_sBlend, bool& x_bToSave, num x_nParaAcel)
  local num l_nSize
  local num l_i
begin
  call getPointSize(x_sKey,l_nSize)
  for l_i = 0 to l_nSize-1
    if trajTemp:tTrajItem[x_sKey].pPointItem[l_i].pParaItem.nMoveType==x_nMoveType
      // trajTemp:tTrajItem[x_sKey].pPointItem[l_i].pParaItem.nMoveType=x_nMoveType
      trajTemp:tTrajItem[x_sKey].pPointItem[l_i].pParaItem.mMdesc.vel=x_nParaSpeed
      trajTemp:tTrajItem[x_sKey].pPointItem[l_i].pParaItem.mMdesc.accel=x_nParaAcel
      trajTemp:tTrajItem[x_sKey].pPointItem[l_i].pParaItem.mMdesc.leave=x_nParaBlend
      trajTemp:tTrajItem[x_sKey].pPointItem[l_i].pParaItem.nPercentage=x_nParaPercent
      switch x_sBlend
        case "OFF"
          trajTemp:tTrajItem[x_sKey].pPointItem[l_i].pParaItem.mMdesc.blend=off
        break
        case "关节"
          trajTemp:tTrajItem[x_sKey].pPointItem[l_i].pParaItem.mMdesc.blend=joint
        break
        case "笛卡尔"
          trajTemp:tTrajItem[x_sKey].pPointItem[l_i].pParaItem.mMdesc.blend=Cartesian
        break
      endSwitch
    endIf
  endFor
  //trajTemp:libSave()
  //delay(0.5)
  logMsg("参数已修改")
  x_bToSave=true
end

--- modifyPara.pgx ---
public program modifyPara(string x_sKey, num x_nIndex, num x_nMoveType, num x_nParaSpeed, num x_nParaBlend, num x_nParaPercent, string x_sComment, bool x_bSafePoint, string x_sBlend, bool& x_bToSave, num& x_nValue[], num x_nParaAcel)
begin
  trajTemp:tTrajItem[x_sKey].pPointItem[x_nIndex].sID=x_sComment
  trajTemp:tTrajItem[x_sKey].pPointItem[x_nIndex].pParaItem.nMoveType=x_nMoveType
  trajTemp:tTrajItem[x_sKey].pPointItem[x_nIndex].pParaItem.mMdesc.vel=x_nParaSpeed
  trajTemp:tTrajItem[x_sKey].pPointItem[x_nIndex].pParaItem.mMdesc.accel=x_nParaAcel
  trajTemp:tTrajItem[x_sKey].pPointItem[x_nIndex].pParaItem.mMdesc.leave=x_nParaBlend
  trajTemp:tTrajItem[x_sKey].pPointItem[x_nIndex].pParaItem.nPercentage=x_nParaPercent
  trajTemp:tTrajItem[x_sKey].pPointItem.pParaItem.bSafePoint=(x_bSafePoint==true)
  switch x_sBlend
    case "OFF"
      trajTemp:tTrajItem[x_sKey].pPointItem[x_nIndex].pParaItem.mMdesc.blend=off
    break
    case "关节"
      trajTemp:tTrajItem[x_sKey].pPointItem[x_nIndex].pParaItem.mMdesc.blend=joint
    break
    case "笛卡尔"
      trajTemp:tTrajItem[x_sKey].pPointItem[x_nIndex].pParaItem.mMdesc.blend=Cartesian
    break

  endSwitch
  switch x_nMoveType
    case 0
      trajTemp:tTrajItem[x_sKey].pPointItem[x_nIndex].jJointRx.j1=x_nValue[0]
      trajTemp:tTrajItem[x_sKey].pPointItem[x_nIndex].jJointRx.j2=x_nValue[1]
      trajTemp:tTrajItem[x_sKey].pPointItem[x_nIndex].jJointRx.j3=x_nValue[2]
      trajTemp:tTrajItem[x_sKey].pPointItem[x_nIndex].jJointRx.j4=x_nValue[3]
      trajTemp:tTrajItem[x_sKey].pPointItem[x_nIndex].jJointRx.j5=x_nValue[4]
      trajTemp:tTrajItem[x_sKey].pPointItem[x_nIndex].jJointRx.j6=x_nValue[5]
    break
    case 1
      trajTemp:tTrajItem[x_sKey].pPointItem[x_nIndex].pPointRx.trsf.x=x_nValue[0]
      trajTemp:tTrajItem[x_sKey].pPointItem[x_nIndex].pPointRx.trsf.y=x_nValue[1]
      trajTemp:tTrajItem[x_sKey].pPointItem[x_nIndex].pPointRx.trsf.z=x_nValue[2]
      trajTemp:tTrajItem[x_sKey].pPointItem[x_nIndex].pPointRx.trsf.rx=x_nValue[3]
      trajTemp:tTrajItem[x_sKey].pPointItem[x_nIndex].pPointRx.trsf.ry=x_nValue[4]
      trajTemp:tTrajItem[x_sKey].pPointItem[x_nIndex].pPointRx.trsf.rz=x_nValue[5]
    break
    case 2
      trajTemp:tTrajItem[x_sKey].pPointItem[x_nIndex].pPointRx.trsf.x=x_nValue[0]
      trajTemp:tTrajItem[x_sKey].pPointItem[x_nIndex].pPointRx.trsf.y=x_nValue[1]
      trajTemp:tTrajItem[x_sKey].pPointItem[x_nIndex].pPointRx.trsf.z=x_nValue[2]
      trajTemp:tTrajItem[x_sKey].pPointItem[x_nIndex].pPointRx.trsf.rx=x_nValue[3]
      trajTemp:tTrajItem[x_sKey].pPointItem[x_nIndex].pPointRx.trsf.ry=x_nValue[4]
      trajTemp:tTrajItem[x_sKey].pPointItem[x_nIndex].pPointRx.trsf.rz=x_nValue[5]
      trajTemp:tTrajItem[x_sKey].pPointItem[x_nIndex].pInter.trsf.x=x_nValue[6]
      trajTemp:tTrajItem[x_sKey].pPointItem[x_nIndex].pInter.trsf.y=x_nValue[7]
      trajTemp:tTrajItem[x_sKey].pPointItem[x_nIndex].pInter.trsf.z=x_nValue[8]
      trajTemp:tTrajItem[x_sKey].pPointItem[x_nIndex].pInter.trsf.rx=x_nValue[9]
      trajTemp:tTrajItem[x_sKey].pPointItem[x_nIndex].pInter.trsf.ry=x_nValue[10]
      trajTemp:tTrajItem[x_sKey].pPointItem[x_nIndex].pInter.trsf.rz=x_nValue[11]
    break
  endSwitch
  //trajTemp:libSave()
  //delay(0.5)
  logMsg("参数已修改")
  x_bToSave=true
end

--- new.pgx ---
public program new(string x_sKey, num x_nFrameIndex, num x_nToolIndex, num x_nMoveID, bool& x_bToSave)
begin
  if !isDefined(trajTemp:tTrajItem[x_sKey]) and x_sKey!=""
    insert(trajTemp:tTrajItem[x_sKey])
    trajTemp:tTrajItem[x_sKey].nFrameIndex=x_nFrameIndex
    trajTemp:tTrajItem[x_sKey].nToolIndex=x_nToolIndex
    trajTemp:tTrajItem[x_sKey].nMoveID=x_nMoveID
    //trajTemp:libSave()
    x_bToSave=true
    delay(0)
  else
    userPageAlert("项目存在，请重新命名！")
  endIf
end

--- onSave.pgx ---
public program onSave(bool& x_bToSave)
begin
  if x_bToSave
    rs:bIsSaving=true
    trajTemp:libSave()
    x_bToSave=false
    rs:bIsSaving=false
    delay(0.5)
    popUpMsg("trajectory数据已保存")
  endIf
end

--- pointEdit.pgx ---
public program pointEdit()
  local bool l_bExit
begin

end

--- pointEditValue.pgx ---
public program pointEditValue(string x_sMoveType, string x_sKey, num x_nIndex, num& x_nTRSF[], string& x_sTRSF[], bool& x_bShow2Point)
begin
  switch x_sMoveType
    case "CIRCLE"
      trajTemp:tTrajItem[x_sKey].pPointItem[x_nIndex].pParaItem.nMoveType=2
      x_nTRSF[0]=trajTemp:tTrajItem[x_sKey].pPointItem[x_nIndex].pPointRx.trsf.x
      x_nTRSF[1]=trajTemp:tTrajItem[x_sKey].pPointItem[x_nIndex].pPointRx.trsf.y
      x_nTRSF[2]=trajTemp:tTrajItem[x_sKey].pPointItem[x_nIndex].pPointRx.trsf.z
      x_nTRSF[3]=trajTemp:tTrajItem[x_sKey].pPointItem[x_nIndex].pPointRx.trsf.rx
      x_nTRSF[4]=trajTemp:tTrajItem[x_sKey].pPointItem[x_nIndex].pPointRx.trsf.ry
      x_nTRSF[5]=trajTemp:tTrajItem[x_sKey].pPointItem[x_nIndex].pPointRx.trsf.rz
      x_nTRSF[6]=trajTemp:tTrajItem[x_sKey].pPointItem[x_nIndex].pInter.trsf.x
      x_nTRSF[7]=trajTemp:tTrajItem[x_sKey].pPointItem[x_nIndex].pInter.trsf.y
      x_nTRSF[8]=trajTemp:tTrajItem[x_sKey].pPointItem[x_nIndex].pInter.trsf.z
      x_nTRSF[9]=trajTemp:tTrajItem[x_sKey].pPointItem[x_nIndex].pInter.trsf.rx
      x_nTRSF[10]=trajTemp:tTrajItem[x_sKey].pPointItem[x_nIndex].pInter.trsf.ry
      x_nTRSF[11]=trajTemp:tTrajItem[x_sKey].pPointItem[x_nIndex].pInter.trsf.rz
      x_sTRSF[0]="X:"
      x_sTRSF[1]="Y:"
      x_sTRSF[2]="Z:"
      x_sTRSF[3]="RX:"
      x_sTRSF[4]="RY:"
      x_sTRSF[5]="RZ:"
      x_sTRSF[6]="2X:"
      x_sTRSF[7]="2Y:"
      x_sTRSF[8]="2Z:"
      x_sTRSF[9]="2RX:"
      x_sTRSF[10]="2RY:"
      x_sTRSF[11]="2RZ:"
      x_bShow2Point=true
    break
    case "POINT"
      trajTemp:tTrajItem[x_sKey].pPointItem[x_nIndex].pParaItem.nMoveType=1
      x_nTRSF[0]=trajTemp:tTrajItem[x_sKey].pPointItem[x_nIndex].pPointRx.trsf.x
      x_nTRSF[1]=trajTemp:tTrajItem[x_sKey].pPointItem[x_nIndex].pPointRx.trsf.y
      x_nTRSF[2]=trajTemp:tTrajItem[x_sKey].pPointItem[x_nIndex].pPointRx.trsf.z
      x_nTRSF[3]=trajTemp:tTrajItem[x_sKey].pPointItem[x_nIndex].pPointRx.trsf.rx
      x_nTRSF[4]=trajTemp:tTrajItem[x_sKey].pPointItem[x_nIndex].pPointRx.trsf.ry
      x_nTRSF[5]=trajTemp:tTrajItem[x_sKey].pPointItem[x_nIndex].pPointRx.trsf.rz
      x_sTRSF[0]="X:"
      x_sTRSF[1]="Y:"
      x_sTRSF[2]="Z:"
      x_sTRSF[3]="RX:"
      x_sTRSF[4]="RY:"
      x_sTRSF[5]="RZ:"
    break
    case "JOINT"
      trajTemp:tTrajItem[x_sKey].pPointItem[x_nIndex].pParaItem.nMoveType=0
      x_nTRSF[0]=trajTemp:tTrajItem[x_sKey].pPointItem[x_nIndex].jJointRx.j1
      x_nTRSF[1]=trajTemp:tTrajItem[x_sKey].pPointItem[x_nIndex].jJointRx.j2
      x_nTRSF[2]=trajTemp:tTrajItem[x_sKey].pPointItem[x_nIndex].jJointRx.j3
      x_nTRSF[3]=trajTemp:tTrajItem[x_sKey].pPointItem[x_nIndex].jJointRx.j4
      x_nTRSF[4]=trajTemp:tTrajItem[x_sKey].pPointItem[x_nIndex].jJointRx.j5
      x_nTRSF[5]=trajTemp:tTrajItem[x_sKey].pPointItem[x_nIndex].jJointRx.j6
      x_sTRSF[0]="J1:"
      x_sTRSF[1]="J2:"
      x_sTRSF[2]="J3:"
      x_sTRSF[3]="J4:"
      x_sTRSF[4]="J5:"
      x_sTRSF[5]="J6:"
    break
  endSwitch
end

--- pointMove.pgx ---
public program pointMove(string x_sKey, num x_nIndex)
  local num l_nType
  local frame l_fFrame
  local pointRx l_pPoint
  local tool l_tTool
  local jointRx l_jJoint
  local bool l_bResult
  local jointRx l_jHere
  local pointRx l_pPoint1
  local num l_nSigIndex
  local bool l_bSigValue
  local num l_nSigValue
  local bool l_bErr
begin
  link(l_fFrame,world)
  link(l_tTool,flange)
  //link(l_pPoint,world)
  l_nType=trajTemp:tTrajItem[x_sKey].pPointItem[x_nIndex].pParaItem.nMoveType
  call savedata:getFrame(trajTemp:tTrajItem[x_sKey].nFrameIndex,l_fFrame)
  call savedata:getTool(trajTemp:tTrajItem[x_sKey].nToolIndex,l_tTool)
  link(l_pPoint,l_fFrame)
  link(l_pPoint1,l_fFrame)
  l_pPoint.trsf=trajTemp:tTrajItem[x_sKey].pPointItem[x_nIndex].pPointRx.trsf
  l_pPoint.config=trajTemp:tTrajItem[x_sKey].pPointItem[x_nIndex].pPointRx.config
  l_pPoint1.trsf=trajTemp:tTrajItem[x_sKey].pPointItem[x_nIndex].pInter.trsf
  l_pPoint1.config=trajTemp:tTrajItem[x_sKey].pPointItem[x_nIndex].pInter.config
  l_jJoint=trajTemp:tTrajItem[x_sKey].pPointItem[x_nIndex].jJointRx
  l_nSigIndex=trajTemp:tTrajItem[x_sKey].pPointItem[x_nIndex].pParaItem.nActionIndex
  l_bSigValue=(trajTemp:tTrajItem[x_sKey].pPointItem[x_nIndex].pParaItem.nSigValue!=0)
  l_nSigValue=trajTemp:tTrajItem[x_sKey].pPointItem[x_nIndex].pParaItem.nSigValue
  if rs:_nOmacStat==9 and workingMode()==1 and isPowered()
    // if !isEmpty()
    stopMove()
    resetMotion()
    l_jHere=herej()
    movej(l_jHere,flange,mSim)
    // endIf
    switch l_nType
      case 1
        call isPointOK(x_sKey,x_nIndex,l_bResult)
        if l_bResult
          movel(l_pPoint,l_tTool,mSim)
        endIf
      break
      case 0
        movej(l_jJoint,l_tTool,mSim)
      break
      case 2
        movec(l_pPoint1,l_pPoint,l_tTool,mSim)
      break
      //Add by Liu Zhengang 20251028
      case 3
        //dIn
        waitEndMove()
        if watch($isKeyPressed(14),5)==true
          call io:waitDigInput(io:dInput[l_nSigIndex],l_bSigValue,l_bErr)
          popUpMsg("din"+"["+toString("",l_nSigIndex)+"]"+"执行成功")
        endIf

      break
      case 4
        //dOut
        waitEndMove()
        if watch($isKeyPressed(14),5)==true

          call io:setDigOutput(io:dOutput[l_nSigIndex],l_bSigValue,l_bErr)
          popUpMsg("dout"+"["+toString("",l_nSigIndex)+"]"+"执行成功")
        endIf
      break
      case 5
        //ain
        waitEndMove()
        if watch($isKeyPressed(14),5)==true
          call io:waitAnaInput(io:aInput[l_nSigIndex],l_nSigValue,l_bErr)
          popUpMsg("ain"+"["+toString("",l_nSigIndex)+"]"+"执行成功")
        endIf

        // wait(l_nSigValue==l_nValue)
      break
      case 6
        //aout
        waitEndMove()
        if watch($isKeyPressed(14),5)==true
          call io:setAnaOutput(io:aOutput[l_nSigIndex],l_nSigValue,l_bErr)
          popUpMsg("aout"+"["+toString("",l_nSigIndex)+"]"+"执行成功")
        endIf
      break
    endSwitch
    delay(0)
  endIf
end

--- pointMove1.pgx ---
public program pointMove1(string x_sKey, num x_nIndex, num x_nPointIndex)
  local num l_nType
  local frame l_fFrame
  local pointRx l_pPoint
  local tool l_tTool
  local jointRx l_jJoint
  local bool l_bResult
  local jointRx l_jHere
begin
  link(l_fFrame,world)
  link(l_tTool,flange)
  //link(l_pPoint,world)
  l_nType=trajTemp:tTrajItem[x_sKey].pPointItem[x_nIndex].pParaItem.nMoveType
  call savedata:getFrame(trajTemp:tTrajItem[x_sKey].nFrameIndex,l_fFrame)
  call savedata:getTool(trajTemp:tTrajItem[x_sKey].nToolIndex,l_tTool)
  link(l_pPoint,l_fFrame)
  switch x_nPointIndex
    case 0
      l_pPoint.trsf=trajTemp:tTrajItem[x_sKey].pPointItem[x_nIndex].pInter.trsf
      l_pPoint.config=trajTemp:tTrajItem[x_sKey].pPointItem[x_nIndex].pInter.config
    break
    case 1
      l_pPoint.trsf=trajTemp:tTrajItem[x_sKey].pPointItem[x_nIndex].pPointRx.trsf
      l_pPoint.config=trajTemp:tTrajItem[x_sKey].pPointItem[x_nIndex].pPointRx.config
    break
  endSwitch

  l_jJoint=trajTemp:tTrajItem[x_sKey].pPointItem[x_nIndex].jJointRx
  if rs:_nOmacStat==9 and workingMode()==1 and isPowered()
    // if !isEmpty()
    stopMove()
    resetMotion()
    l_jHere=herej()
    movej(l_jHere,flange,mSim)
    // endIf
    //    switch l_nType
    //      case 1
    call isPointOK(x_sKey,x_nIndex,l_bResult)
    if l_bResult
      //          movel(l_pPoint,l_tTool,mSim)
      //        endIf
      //      break
      //      case 0
      movej(l_pPoint,l_tTool,mSim)
      waitEndMove()
    endIf
    //      break
    //    endSwitch
    delay(0)
  endIf
end

--- pointToString.pgx ---
public program pointToString(string& x_sMsg, string x_sKey, num x_nIndex)
  local trsf l_trsf
  local string l_sMsg
  local num l_nType
  local jointRx l_jJoint
  local num l_nActionIndex
  local num l_nSigValue
  local num l_nSigType[3]
  local num l_nSigIndex[3]
  local num l_nValue[3]
  local string l_sType[3]
  local string l_sValue[3]
  local num l_nANDOR[2]
  local string l_sANDOR[2]
  local string l_sSigIndex[3]
  local num l_i
  local num l_nSpeed
  local mdesc l_mdesc
  local string l_sblend
  local string l_sComment
  local bool l_bSafePoint
  local num l_nIndex
  local bool l_bNull[3]
  local bool l_bMark
  local trsf l_trsf1
  local bool l_bErr
begin
  l_nType=trajTemp:tTrajItem[x_sKey].pPointItem[x_nIndex].pParaItem.nMoveType
  l_bMark=(trajTemp:tTrajItem[x_sKey].pPointItem[x_nIndex].bMarked==true)
  switch l_nType
    //关节
    case 0
      l_jJoint=trajTemp:tTrajItem[x_sKey].pPointItem[x_nIndex].jJointRx
      l_mdesc=trajTemp:tTrajItem[x_sKey].pPointItem[x_nIndex].pParaItem.mMdesc
      l_sComment=trajTemp:tTrajItem[x_sKey].pPointItem[x_nIndex].sID
      l_bSafePoint=(trajTemp:tTrajItem[x_sKey].pPointItem[x_nIndex].pParaItem.bSafePoint==true)
      if l_mdesc.blend!=off
        l_sblend=toString("",l_mdesc.leave)
      else
        l_sblend="off"
      endIf
      l_sMsg=", J["
      l_sMsg=l_sMsg+toString("",l_jJoint.j1)+", "
      l_sMsg=l_sMsg+toString("",l_jJoint.j2)+", "
      l_sMsg=l_sMsg+toString("",l_jJoint.j3)+", "
      l_sMsg=l_sMsg+toString("",l_jJoint.j4)+", "
      l_sMsg=l_sMsg+toString("",l_jJoint.j5)+", "
      l_sMsg=l_sMsg+toString("",l_jJoint.j6)+"]"
      l_sMsg=l_sMsg+"_spd="+toString("",l_mdesc.vel)+"%"
      l_sMsg=l_sMsg+"_b="+l_sblend
      if l_bSafePoint
        l_sMsg=l_sMsg+" @safepoint"
      endIf
      if l_sComment!=""
        l_sMsg=l_sMsg+"#"+l_sComment
      endIf
    break
    //
    case 1
      l_bSafePoint=(trajTemp:tTrajItem[x_sKey].pPointItem[x_nIndex].pParaItem.bSafePoint==true)
      l_trsf=trajTemp:tTrajItem[x_sKey].pPointItem[x_nIndex].pPointRx.trsf
      l_mdesc=trajTemp:tTrajItem[x_sKey].pPointItem[x_nIndex].pParaItem.mMdesc
      l_sComment=trajTemp:tTrajItem[x_sKey].pPointItem[x_nIndex].sID
      if l_mdesc.blend!=off
        l_sblend=toString("",l_mdesc.leave)
      else
        l_sblend="off"
      endIf
      l_sMsg=", L["
      l_sMsg=l_sMsg+toString("",l_trsf.x)+","
      l_sMsg=l_sMsg+toString("",l_trsf.y)+","
      l_sMsg=l_sMsg+toString("",l_trsf.z)+","
      l_sMsg=l_sMsg+toString("",l_trsf.rx)+","
      l_sMsg=l_sMsg+toString("",l_trsf.ry)+","
      l_sMsg=l_sMsg+toString("",l_trsf.rz)+"]"
      l_sMsg=l_sMsg+"_spd="+toString("",l_mdesc.vel)+"%"
      l_sMsg=l_sMsg+"_b="+l_sblend
      if l_bSafePoint
        l_sMsg=l_sMsg+"_@safepoint"
      endIf
      if l_sComment!=""
        l_sMsg=l_sMsg+ "#"+l_sComment+""
      endIf

    break
    //2024.12.23 add圆弧
    case 2
      l_bSafePoint=(trajTemp:tTrajItem[x_sKey].pPointItem[x_nIndex].pParaItem.bSafePoint==true)
      l_trsf=trajTemp:tTrajItem[x_sKey].pPointItem[x_nIndex].pPointRx.trsf
      l_trsf1=trajTemp:tTrajItem[x_sKey].pPointItem[x_nIndex].pInter.trsf
      l_mdesc=trajTemp:tTrajItem[x_sKey].pPointItem[x_nIndex].pParaItem.mMdesc
      l_sComment=trajTemp:tTrajItem[x_sKey].pPointItem[x_nIndex].sID
      if l_mdesc.blend!=off
        l_sblend=toString("",l_mdesc.leave)
      else
        l_sblend="off"
      endIf
      l_sMsg=", C["
      l_sMsg=l_sMsg+toString("",l_trsf.x)+","
      l_sMsg=l_sMsg+toString("",l_trsf.y)+","
      l_sMsg=l_sMsg+toString("",l_trsf.z)+","
      l_sMsg=l_sMsg+toString("",l_trsf.rx)+","
      l_sMsg=l_sMsg+toString("",l_trsf.ry)+","
      l_sMsg=l_sMsg+toString("",l_trsf.rz)+"]["
      l_sMsg=l_sMsg+toString("",l_trsf1.x)+","
      l_sMsg=l_sMsg+toString("",l_trsf1.y)+","
      l_sMsg=l_sMsg+toString("",l_trsf1.z)+","
      l_sMsg=l_sMsg+toString("",l_trsf1.rx)+","
      l_sMsg=l_sMsg+toString("",l_trsf1.ry)+","
      l_sMsg=l_sMsg+toString("",l_trsf1.rz)+"]"
      l_sMsg=l_sMsg+"_spd="+toString("",l_mdesc.vel)+"%"
      l_sMsg=l_sMsg+"_b="+l_sblend
      if l_bSafePoint
        l_sMsg=l_sMsg+"_@safepoint"
      endIf
      if l_sComment!=""
        l_sMsg=l_sMsg+ "#"+l_sComment+""
      endIf
    break
    case 3
      l_sMsg=", wait->DIN["
      l_nActionIndex=trajTemp:tTrajItem[x_sKey].pPointItem[x_nIndex].pParaItem.nActionIndex
      l_nSigValue=trajTemp:tTrajItem[x_sKey].pPointItem[x_nIndex].pParaItem.nSigValue
      l_sMsg=l_sMsg+toString("",l_nActionIndex)+"]-"+io:dInItem[l_nActionIndex].sComment+"="
      if l_nSigValue!=0
        l_sMsg=l_sMsg+"TRUE"
      else
        l_sMsg=l_sMsg+"FALSE"
      endIf
    break
    case 4
      l_sMsg=", DOUT["
      l_nActionIndex=trajTemp:tTrajItem[x_sKey].pPointItem[x_nIndex].pParaItem.nActionIndex
      l_nSigValue=trajTemp:tTrajItem[x_sKey].pPointItem[x_nIndex].pParaItem.nSigValue
      l_sMsg=l_sMsg+toString("",l_nActionIndex)+"]-"+io:dOutItem[l_nActionIndex].sComment+"="
      if l_nSigValue!=0
        l_sMsg=l_sMsg+"TRUE"
      else
        l_sMsg=l_sMsg+"FALSE"
      endIf
    break
    case 5
      l_sMsg=", wait->AIN["
      l_nActionIndex=trajTemp:tTrajItem[x_sKey].pPointItem[x_nIndex].pParaItem.nActionIndex
      l_nSigValue=trajTemp:tTrajItem[x_sKey].pPointItem[x_nIndex].pParaItem.nSigValue
      l_sMsg=l_sMsg+toString("",l_nActionIndex)+"]-"+io:aInItem[l_nActionIndex].sComment+"="
      l_sMsg=l_sMsg+toString(".3",l_nSigValue)
    break
    case 6
      l_sMsg=", AOUT["
      l_nActionIndex=trajTemp:tTrajItem[x_sKey].pPointItem[x_nIndex].pParaItem.nActionIndex
      l_nSigValue=trajTemp:tTrajItem[x_sKey].pPointItem[x_nIndex].pParaItem.nSigValue
      l_sMsg=l_sMsg+toString("",l_nActionIndex)+"]-"+io:aOutItem[l_nActionIndex].sComment+"="
      l_sMsg=l_sMsg+toString(".3",l_nSigValue)
    break
    case 7
      l_sMsg=", DELAY = "
      l_nSigValue=trajTemp:tTrajItem[x_sKey].pPointItem[x_nIndex].pParaItem.nDelay
      l_sMsg=l_sMsg+toString(".3",l_nSigValue)+" s"
    break
    case 8
      l_sMsg=", IF "
      for l_i = 0 to 2
        l_bNull[l_i]=true
        l_nSigType[l_i]=trajTemp:tTrajItem[x_sKey].pPointItem[x_nIndex].pParaItem.iIfItem.nSigType[l_i]
        l_nValue[l_i]=trajTemp:tTrajItem[x_sKey].pPointItem[x_nIndex].pParaItem.iIfItem.nValue[l_i]
        l_nSigIndex[l_i]=trajTemp:tTrajItem[x_sKey].pPointItem[x_nIndex].pParaItem.iIfItem.nSigIndex[l_i]
        l_sSigIndex[l_i]=toString("",l_nSigIndex[l_i])
        switch l_nSigType[l_i]
          case 1
            l_sType[l_i]="DIN"
            if l_nValue[l_i]!=0
              l_sValue[l_i]="TRUE"
            else
              l_sValue[l_i]="FALSE"
            endIf
          break
          case 2
            l_sType[l_i]="DOUT"
            if l_nValue[l_i]!=0
              l_sValue[l_i]="TRUE"
            else
              l_sValue[l_i]="FALSE"
            endIf
          break
          case 3
            l_sType[l_i]="AIN"
            l_sValue[l_i]=toString(".2",l_nValue[l_i])
          break
          case 4
            l_sType[l_i]="AOUT"
            l_sValue[l_i]=toString(".2",l_nValue[l_i])
          break
          default
            l_bNull[l_i]=false
          break
        endSwitch

      endFor
      for l_i = 0 to 1
        if trajTemp:tTrajItem[x_sKey].pPointItem[x_nIndex].pParaItem.iIfItem.bANDOR[l_i]
          l_sANDOR[l_i]="or"
        else
          l_sANDOR[l_i]="and"
        endIf
      endFor
      //l_sMsg=""
      if l_bNull[0] and l_bNull[1] and l_bNull[2]
        l_sMsg=l_sMsg+l_sType[0]+"["+l_sSigIndex[0]+"]="+l_sValue[0] +" "+l_sANDOR[0]+" "
        l_sMsg=l_sMsg+l_sType[1]+"["+l_sSigIndex[1]+"]="+l_sValue[1] +" "+l_sANDOR[1]+" "
        l_sMsg=l_sMsg+l_sType[2]+"["+l_sSigIndex[2]+"]="+l_sValue[2]
      elseIf l_bNull[0] and !l_bNull[1] and !l_bNull[2]
        l_sMsg=l_sMsg+l_sType[0]+"["+l_sSigIndex[0]+"]="+l_sValue[0]
      elseIf l_bNull[0] and l_bNull[1] and !l_bNull[2]
        l_sMsg=l_sMsg+l_sType[0]+"["+l_sSigIndex[0]+"]="+l_sValue[0] +" "+l_sANDOR[0]+" "
        l_sMsg=l_sMsg+l_sType[1]+"["+l_sSigIndex[1]+"]="+l_sValue[1]
      elseIf !l_bNull[0] and l_bNull[1] and !l_bNull[2]
        l_sMsg=l_sMsg+l_sType[1]+"["+l_sSigIndex[1]+"]="+l_sValue[1]
      elseIf !l_bNull[0] and !l_bNull[1] and l_bNull[2]
        l_sMsg=l_sMsg+l_sType[2]+"["+l_sSigIndex[2]+"]="+l_sValue[2]
      elseIf l_bNull[0] and !l_bNull[1] and l_bNull[2]
        l_sMsg=l_sMsg+l_sType[0]+"["+l_sSigIndex[0]+"]="+l_sValue[0] +" "+l_sANDOR[0]+" "
        l_sMsg=l_sMsg+l_sType[2]+"["+l_sSigIndex[2]+"]="+l_sValue[2]
      elseIf !l_bNull[0] and l_bNull[1] and l_bNull[2]
        l_sMsg=l_sMsg+l_sType[1]+"["+l_sSigIndex[1]+"]="+l_sValue[1] +" "+l_sANDOR[1]+" "
        l_sMsg=l_sMsg+l_sType[2]+"["+l_sSigIndex[2]+"]="+l_sValue[2]
      endIf
    break
    case 9
      l_sMsg=",  ENDIF"
    break
    case 10
      //action
      l_nIndex=trajTemp:tTrajItem[x_sKey].pPointItem[x_nIndex].pParaItem.nSigValue
      l_sComment=actData:aActItem[l_nIndex].sComment
      l_sMsg=",Action:"+l_sComment
    break
    case 11
      //2025.7.21 add 喷淋delay
      l_sMsg=", WASH_DELAY = "
      call io:getAnaIO(io:aInput[15],l_nSigValue,l_bErr)
      l_sMsg=l_sMsg+toString(".3",l_nSigValue)+" s"
    break
  endSwitch
  //是否被标记
  if l_bMark
    l_sMsg=",*,"+l_sMsg
  endIf


  x_sMsg=l_sMsg
end

--- resetMark.pgx ---
public program resetMark(string x_sKey)
  local num l_nSize
  local num l_i
begin
  call getPointSize(x_sKey,l_nSize)
  //resize(savedata:nMarkIndex,1,l_nSize)
  for l_i = 0 to l_nSize-1
    trajTemp:tTrajItem[x_sKey].pPointItem[l_i].bMarked=false
  endFor
end

--- resizeMark.pgx ---
public program resizeMark(string x_sKey)
  local num l_nSize
  local num l_i
begin
  call getPointSize(x_sKey,l_nSize)
  //resize(savedata:nMarkIndex,1,l_nSize)
  for l_i = 0 to l_nSize-1
    trajTemp:tTrajItem[x_sKey].pPointItem[l_i].bMarked=false
  endFor
end

--- setMark.pgx ---
public program setMark(string x_sKey, num x_nIndex)
begin

  trajTemp:tTrajItem[x_sKey].pPointItem[x_nIndex].bMarked=!trajTemp:tTrajItem[x_sKey].pPointItem[x_nIndex].bMarked
//  if trajTemp:tTrajItem[x_sKey].pPointItem[x_nIndex].bMarked
//    savedata:nMarkIndex[x_nIndex]=1
//  else
//    savedata:nMarkIndex[x_nIndex]=-1
//  endIf

end

--- stop.pgx ---
program stop()
begin
end

--- teachPoint.pgx ---
public program teachPoint(string x_sKey, num x_nIndex, bool& x_bToSave)
  local num l_nFrameIndex
  local num l_nToolIndex
  local frame l_fFrame
  local tool l_tTool
  local bool l_bResult
  local pointRx l_pPoint
begin
  link(l_tTool,flange)
  link(l_fFrame,world)
  l_bResult=userPageConfirm("是否记录当前点位："+toString("",x_nIndex))
  if l_bResult
    l_nFrameIndex=trajTemp:tTrajItem[x_sKey].nFrameIndex
    l_nToolIndex=trajTemp:tTrajItem[x_sKey].nToolIndex
    call savedata:getFrame(l_nFrameIndex,l_fFrame)
    call savedata:getTool(l_nToolIndex,l_tTool)


    trajTemp:tTrajItem[x_sKey].pPointItem[x_nIndex].jJointRx=herej()
    l_pPoint=jointToPoint(l_tTool,l_fFrame,herej())
    trajTemp:tTrajItem[x_sKey].pPointItem[x_nIndex].pPointRx.trsf=l_pPoint.trsf
    trajTemp:tTrajItem[x_sKey].pPointItem[x_nIndex].pPointRx.config=l_pPoint.config
    x_bToSave=true
  endIf
end

--- teachPoint1.pgx ---
public program teachPoint1(string x_sKey, num x_nIndex, num x_nPointIndex)
  local num l_nFrameIndex
  local num l_nToolIndex
  local frame l_fFrame
  local tool l_tTool
  local bool l_bResult
  local pointRx l_pPoint
begin
  link(l_tTool,flange)
  link(l_fFrame,world)
  //  l_bResult=userPageConfirm("是否记录当前点位："+toString("",x_nIndex))
  //  if l_bResult
  l_nFrameIndex=trajTemp:tTrajItem[x_sKey].nFrameIndex
  l_nToolIndex=trajTemp:tTrajItem[x_sKey].nToolIndex
  call savedata:getFrame(l_nFrameIndex,l_fFrame)
  call savedata:getTool(l_nToolIndex,l_tTool)


  trajTemp:tTrajItem[x_sKey].pPointItem[x_nIndex].jJointRx=herej()
  l_pPoint=jointToPoint(l_tTool,l_fFrame,herej())
  switch x_nPointIndex
    case 0
      trajTemp:tTrajItem[x_sKey].pPointItem[x_nIndex].pInter.trsf=l_pPoint.trsf
      trajTemp:tTrajItem[x_sKey].pPointItem[x_nIndex].pInter.config=l_pPoint.config
    break
    case 1
      trajTemp:tTrajItem[x_sKey].pPointItem[x_nIndex].pPointRx.trsf=l_pPoint.trsf
      trajTemp:tTrajItem[x_sKey].pPointItem[x_nIndex].pPointRx.config=l_pPoint.config
    break
  endSwitch

  //x_bToSave=true
  //  endIf
end
